FUNCTION_BLOCK MGE_Generico_HMI (* Service Interface Function Block Type *)
  (* Standard: 61499-2 *)
  (* Version 1.5, 15/10/2026, Hidryco, Hidryco, IHM do MGE_Generico (tags do MGE antigo mantidas) *)
  PACKAGE Hidryco.HidrycoLib;
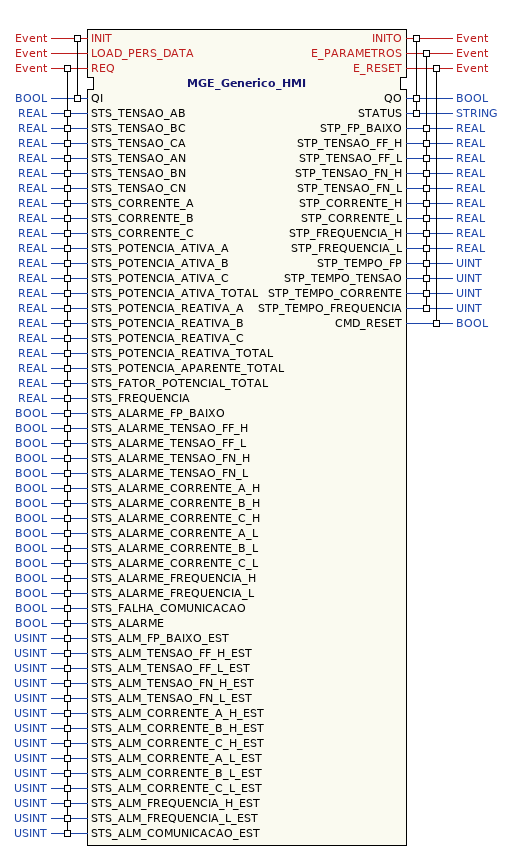
  EVENT_INPUT
    INIT WITH QI;
    LOAD_PERS_DATA; (* Reenvia os parametros persistentes *)
    REQ WITH STS_TENSAO_AB, STS_TENSAO_BC, STS_TENSAO_CA, STS_TENSAO_AN, STS_TENSAO_BN, STS_TENSAO_CN, STS_CORRENTE_A, STS_CORRENTE_B, STS_CORRENTE_C, STS_POTENCIA_ATIVA_A, STS_POTENCIA_ATIVA_B, STS_POTENCIA_ATIVA_C, STS_POTENCIA_ATIVA_TOTAL, STS_POTENCIA_REATIVA_A, STS_POTENCIA_REATIVA_B, STS_POTENCIA_REATIVA_C, STS_POTENCIA_REATIVA_TOTAL, STS_POTENCIA_APARENTE_TOTAL, STS_FATOR_POTENCIAL_TOTAL, STS_FREQUENCIA, STS_ALARME_FP_BAIXO, STS_ALARME_TENSAO_FF_H, STS_ALARME_TENSAO_FF_L, STS_ALARME_TENSAO_FN_H, STS_ALARME_TENSAO_FN_L, STS_ALARME_CORRENTE_A_H, STS_ALARME_CORRENTE_B_H, STS_ALARME_CORRENTE_C_H, STS_ALARME_CORRENTE_A_L, STS_ALARME_CORRENTE_B_L, STS_ALARME_CORRENTE_C_L, STS_ALARME_FREQUENCIA_H, STS_ALARME_FREQUENCIA_L, STS_FALHA_COMUNICACAO, STS_ALARME, STS_ALM_FP_BAIXO_EST, STS_ALM_TENSAO_FF_H_EST, STS_ALM_TENSAO_FF_L_EST, STS_ALM_TENSAO_FN_H_EST, STS_ALM_TENSAO_FN_L_EST, STS_ALM_CORRENTE_A_H_EST, STS_ALM_CORRENTE_B_H_EST, STS_ALM_CORRENTE_C_H_EST, STS_ALM_CORRENTE_A_L_EST, STS_ALM_CORRENTE_B_L_EST, STS_ALM_CORRENTE_C_L_EST, STS_ALM_FREQUENCIA_H_EST, STS_ALM_FREQUENCIA_L_EST, STS_ALM_COMUNICACAO_EST; (* Atualizacao de status *)
  END_EVENT
  EVENT_OUTPUT
    INITO WITH QO, STATUS;
    E_PARAMETROS WITH STP_FP_BAIXO, STP_TENSAO_FF_H, STP_TENSAO_FF_L, STP_TENSAO_FN_H, STP_TENSAO_FN_L, STP_CORRENTE_H, STP_CORRENTE_L, STP_FREQUENCIA_H, STP_FREQUENCIA_L, STP_TEMPO_FP, STP_TEMPO_TENSAO, STP_TEMPO_CORRENTE, STP_TEMPO_FREQUENCIA;
    E_RESET WITH CMD_RESET;
  END_EVENT
  VAR_INPUT
    QI : BOOL;
    STS_TENSAO_AB : REAL; (* Tensao A-B (V) *)
    STS_TENSAO_BC : REAL; (* Tensao B-C (V) *)
    STS_TENSAO_CA : REAL; (* Tensao C-A (V) *)
    STS_TENSAO_AN : REAL; (* Tensao A-N (V) *)
    STS_TENSAO_BN : REAL; (* Tensao B-N (V) *)
    STS_TENSAO_CN : REAL; (* Tensao C-N (V) *)
    STS_CORRENTE_A : REAL; (* Corrente fase A (A) *)
    STS_CORRENTE_B : REAL; (* Corrente fase B (A) *)
    STS_CORRENTE_C : REAL; (* Corrente fase C (A) *)
    STS_POTENCIA_ATIVA_A : REAL; (* Potencia ativa fase A (kW) *)
    STS_POTENCIA_ATIVA_B : REAL; (* Potencia ativa fase B (kW) *)
    STS_POTENCIA_ATIVA_C : REAL; (* Potencia ativa fase C (kW) *)
    STS_POTENCIA_ATIVA_TOTAL : REAL; (* Potencia ativa total (kW) *)
    STS_POTENCIA_REATIVA_A : REAL; (* Potencia reativa fase A (kVAr) *)
    STS_POTENCIA_REATIVA_B : REAL; (* Potencia reativa fase B (kVAr) *)
    STS_POTENCIA_REATIVA_C : REAL; (* Potencia reativa fase C (kVAr) *)
    STS_POTENCIA_REATIVA_TOTAL : REAL; (* Potencia reativa total (kVAr) *)
    STS_POTENCIA_APARENTE_TOTAL : REAL; (* Potencia aparente total (kVA) *)
    STS_FATOR_POTENCIAL_TOTAL : REAL; (* Fator de potencia total *)
    STS_FREQUENCIA : REAL; (* Frequencia (Hz) *)
    STS_ALARME_FP_BAIXO : BOOL; (* Fator de potência baixo *)
    STS_ALARME_TENSAO_FF_H : BOOL; (* Tensão entre fases alta *)
    STS_ALARME_TENSAO_FF_L : BOOL; (* Tensão entre fases baixa *)
    STS_ALARME_TENSAO_FN_H : BOOL; (* Tensão fase-neutro alta *)
    STS_ALARME_TENSAO_FN_L : BOOL; (* Tensão fase-neutro baixa *)
    STS_ALARME_CORRENTE_A_H : BOOL; (* Corrente fase A alta *)
    STS_ALARME_CORRENTE_B_H : BOOL; (* Corrente fase B alta *)
    STS_ALARME_CORRENTE_C_H : BOOL; (* Corrente fase C alta *)
    STS_ALARME_CORRENTE_A_L : BOOL; (* Corrente fase A baixa *)
    STS_ALARME_CORRENTE_B_L : BOOL; (* Corrente fase B baixa *)
    STS_ALARME_CORRENTE_C_L : BOOL; (* Corrente fase C baixa *)
    STS_ALARME_FREQUENCIA_H : BOOL; (* Frequência alta *)
    STS_ALARME_FREQUENCIA_L : BOOL; (* Frequência baixa *)
    STS_FALHA_COMUNICACAO : BOOL; (* Falha de comunicacao *)
    STS_ALARME : BOOL; (* Algum alarme do medidor *)
    STS_ALM_FP_BAIXO_EST : USINT; (* Estado do ALARM_BIT Fator de potência baixo (0 normal, 1 ativo reconhecido, 2 ativo nao reconhecido, 3 saiu nao reconhecido, 4 ativo e saiu nao reconhecido) *)
    STS_ALM_TENSAO_FF_H_EST : USINT; (* Estado do ALARM_BIT Tensão entre fases alta (0 normal, 1 ativo reconhecido, 2 ativo nao reconhecido, 3 saiu nao reconhecido, 4 ativo e saiu nao reconhecido) *)
    STS_ALM_TENSAO_FF_L_EST : USINT; (* Estado do ALARM_BIT Tensão entre fases baixa (0 normal, 1 ativo reconhecido, 2 ativo nao reconhecido, 3 saiu nao reconhecido, 4 ativo e saiu nao reconhecido) *)
    STS_ALM_TENSAO_FN_H_EST : USINT; (* Estado do ALARM_BIT Tensão fase-neutro alta (0 normal, 1 ativo reconhecido, 2 ativo nao reconhecido, 3 saiu nao reconhecido, 4 ativo e saiu nao reconhecido) *)
    STS_ALM_TENSAO_FN_L_EST : USINT; (* Estado do ALARM_BIT Tensão fase-neutro baixa (0 normal, 1 ativo reconhecido, 2 ativo nao reconhecido, 3 saiu nao reconhecido, 4 ativo e saiu nao reconhecido) *)
    STS_ALM_CORRENTE_A_H_EST : USINT; (* Estado do ALARM_BIT Corrente fase A alta (0 normal, 1 ativo reconhecido, 2 ativo nao reconhecido, 3 saiu nao reconhecido, 4 ativo e saiu nao reconhecido) *)
    STS_ALM_CORRENTE_B_H_EST : USINT; (* Estado do ALARM_BIT Corrente fase B alta (0 normal, 1 ativo reconhecido, 2 ativo nao reconhecido, 3 saiu nao reconhecido, 4 ativo e saiu nao reconhecido) *)
    STS_ALM_CORRENTE_C_H_EST : USINT; (* Estado do ALARM_BIT Corrente fase C alta (0 normal, 1 ativo reconhecido, 2 ativo nao reconhecido, 3 saiu nao reconhecido, 4 ativo e saiu nao reconhecido) *)
    STS_ALM_CORRENTE_A_L_EST : USINT; (* Estado do ALARM_BIT Corrente fase A baixa (0 normal, 1 ativo reconhecido, 2 ativo nao reconhecido, 3 saiu nao reconhecido, 4 ativo e saiu nao reconhecido) *)
    STS_ALM_CORRENTE_B_L_EST : USINT; (* Estado do ALARM_BIT Corrente fase B baixa (0 normal, 1 ativo reconhecido, 2 ativo nao reconhecido, 3 saiu nao reconhecido, 4 ativo e saiu nao reconhecido) *)
    STS_ALM_CORRENTE_C_L_EST : USINT; (* Estado do ALARM_BIT Corrente fase C baixa (0 normal, 1 ativo reconhecido, 2 ativo nao reconhecido, 3 saiu nao reconhecido, 4 ativo e saiu nao reconhecido) *)
    STS_ALM_FREQUENCIA_H_EST : USINT; (* Estado do ALARM_BIT Frequência alta (0 normal, 1 ativo reconhecido, 2 ativo nao reconhecido, 3 saiu nao reconhecido, 4 ativo e saiu nao reconhecido) *)
    STS_ALM_FREQUENCIA_L_EST : USINT; (* Estado do ALARM_BIT Frequência baixa (0 normal, 1 ativo reconhecido, 2 ativo nao reconhecido, 3 saiu nao reconhecido, 4 ativo e saiu nao reconhecido) *)
    STS_ALM_COMUNICACAO_EST : USINT; (* Estado do ALARM_BIT falha de comunicacao (0 normal, 1 ativo reconhecido, 2 ativo nao reconhecido, 3 saiu nao reconhecido, 4 ativo e saiu nao reconhecido) *)
  END_VAR
  VAR_OUTPUT
    QO : BOOL; (* Event Output Qualifier *)
    STATUS : STRING; (* Service Status *)
    STP_FP_BAIXO : REAL; (* Fator de potência baixo (abaixo de): valor de referencia (adimensional; 0 = desligado) *)
    STP_TENSAO_FF_H : REAL; (* Tensão entre fases alta (acima de): valor de referencia (V; 0 = desligado) *)
    STP_TENSAO_FF_L : REAL; (* Tensão entre fases baixa (abaixo de): valor de referencia (V; 0 = desligado) *)
    STP_TENSAO_FN_H : REAL; (* Tensão fase-neutro alta (acima de): valor de referencia (V; 0 = desligado) *)
    STP_TENSAO_FN_L : REAL; (* Tensão fase-neutro baixa (abaixo de): valor de referencia (V; 0 = desligado) *)
    STP_CORRENTE_H : REAL; (* Corrente alta - fases A, B e C (acima de): valor de referencia (A; 0 = desligado) *)
    STP_CORRENTE_L : REAL; (* Corrente baixa - fases A, B e C (abaixo de): valor de referencia (A; 0 = desligado) *)
    STP_FREQUENCIA_H : REAL; (* Frequência alta (acima de): valor de referencia (Hz; 0 = desligado) *)
    STP_FREQUENCIA_L : REAL; (* Frequência baixa (abaixo de): valor de referencia (Hz; 0 = desligado) *)
    STP_TEMPO_FP : UINT; (* Tempo de retardo (s) dos alarmes de fator de potência *)
    STP_TEMPO_TENSAO : UINT; (* Tempo de retardo (s) dos alarmes de tensão *)
    STP_TEMPO_CORRENTE : UINT; (* Tempo de retardo (s) dos alarmes de corrente *)
    STP_TEMPO_FREQUENCIA : UINT; (* Tempo de retardo (s) dos alarmes de frequência *)
    CMD_RESET : BOOL; (* Reconhece e faz o reset dos alarmes do medidor *)
  END_VAR
  SERVICE /
    SEQUENCE 
    END_SEQUENCE
  END_SERVICE
END_FUNCTION_BLOCK
